# EPICS autosave request: iocs/ad/mythen-ioc/auto_settings.req
file "ADBase_settings.req",         P=$(P),  R=cam1:
$(P)cam1:AcquireTime.PREC
# C includes NDFile_settings.req for cam1:, which mythen.template lacks.
file "mythen_settings.req",       P=$(P),  R=cam1:
file "NDPluginBase_settings.req",   P=$(P),  R=image1:
file "NDStdArrays_settings.req",    P=$(P),  R=image1:
file "commonPlugin_settings.req",   P=$(P)
